PROGRAM main
  VAR
    Water_Level AT %MD0 : REAL := 0.0;
    Low_Level : BOOL;
    High_Level : BOOL;
    Pump AT %QX0.0 : BOOL;
  END_VAR

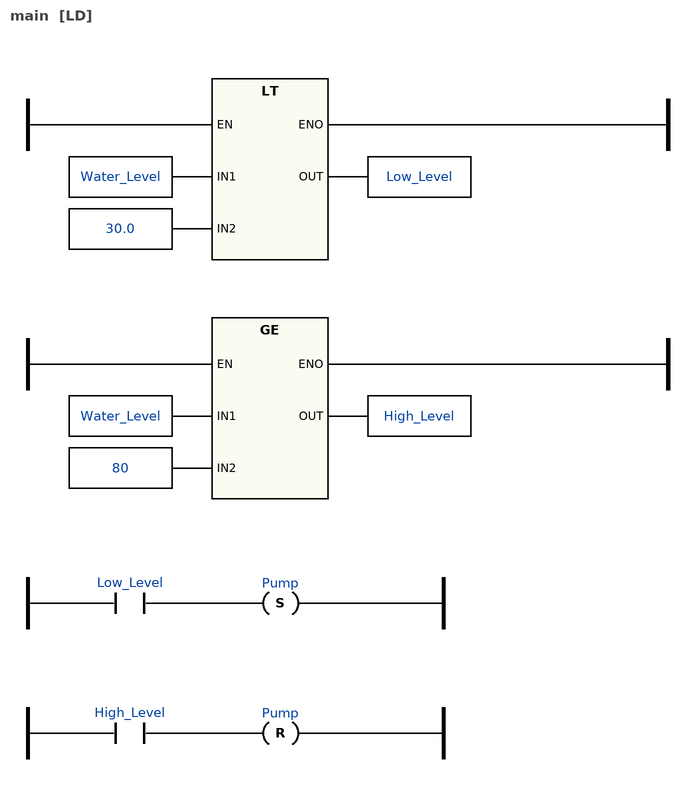
(* LD diagram, written out as Structured Text *)
Low_Level := Water_Level < 30.0;
High_Level := Water_Level >= 80;
IF Low_Level THEN Pump := TRUE; END_IF;
IF High_Level THEN Pump := FALSE; END_IF;
END_PROGRAM
